(* IEC 61131-3 sources: volt/packages/volt-lsp-iec/test-corpus/pro2193/Device/Plc Logic/Application/09 Misc/Library Manager/CAA SegBufMan, 38 files *)

(* ---- ERROR.dut ---- *)
TYPE ERROR :
(
	NO_ERROR := 0,
	FIRST_ERROR := 6100,
	TIME_OUT,
	FIRST_MF,
	LAST_ERROR := 6199
);
END_TYPE

(* ---- RSHANDLING.gvl ---- *)
VAR_GLOBAL
	G_BUFFERCLASS : BufferClass;
	G_QUEUECLASS : QueueClass;
END_VAR

(* ---- VERSIONCONSTANTS.gvl ---- *)
VAR_GLOBAL
	GC_BYVERSION : BYTE := 1;
	GC_BYVERSION_1 : BYTE := 0;
END_VAR

(* ---- _BUFFERADDREF.pou ---- *)
FUNCTION _BUFFERADDREF : ERROR
VAR_INPUT
	HBUFFER : CAA.HANDLE;
END_VAR
END_FUNCTION

(* ---- _CHAINBUFFER.pou ---- *)
FUNCTION _CHAINBUFFER : CAA.HANDLE
VAR_INPUT
	HHEAD : CAA.HANDLE;
	HTAIL : CAA.HANDLE;
	PEERROR : POINTER TO ERROR;
END_VAR
END_FUNCTION

(* ---- _COPYBUFFERDATA.pou ---- *)
FUNCTION _COPYBUFFERDATA : ERROR
VAR_INPUT
	HBUFFER : CAA.HANDLE;
	SZOFFSET : CAA.SIZE;
	SZLENGTH : CAA.SIZE;
	PDATA : CAA.PVOID;
	SZSIZE : CAA.SIZE;
END_VAR
END_FUNCTION

(* ---- _CREATEBUFFER.pou ---- *)
FUNCTION _CREATEBUFFER : CAA.HANDLE
VAR_INPUT
	SZSIZE : CAA.SIZE;
	PDATA : CAA.PVOID;
	XPERMANENT : BOOL;
	PEERROR : POINTER TO ERROR;
END_VAR
END_FUNCTION

(* ---- _CREATEQUEUE.pou ---- *)
FUNCTION _CREATEQUEUE : CAA.HANDLE
VAR_INPUT
	PEERROR : POINTER TO ERROR;
END_VAR
END_FUNCTION

(* ---- _DELETEBUFFER.pou ---- *)
FUNCTION _DELETEBUFFER : ERROR
VAR_INPUT
	HBUFFER : CAA.HANDLE;
END_VAR
END_FUNCTION

(* ---- _DELETEQUEUE.pou ---- *)
FUNCTION _DELETEQUEUE : ERROR
VAR_INPUT
	HQUEUE : CAA.HANDLE;
END_VAR
END_FUNCTION

(* ---- _DEQUEUEBUFFER.pou ---- *)
FUNCTION _DEQUEUEBUFFER : CAA.HANDLE
VAR_INPUT
	HQUEUE : CAA.HANDLE;
	PEERROR : POINTER TO ERROR;
END_VAR
END_FUNCTION

(* ---- _ENQUEUEBUFFER.pou ---- *)
FUNCTION _ENQUEUEBUFFER : ERROR
VAR_INPUT
	HQUEUE : CAA.HANDLE;
	HBUFFER : CAA.HANDLE;
END_VAR
END_FUNCTION

(* ---- _GETBUFFERSIZE.pou ---- *)
FUNCTION _GETBUFFERSIZE : CAA.SIZE
VAR_INPUT
	HBUFFER : CAA.HANDLE;
	PEERROR : POINTER TO ERROR;
END_VAR
END_FUNCTION

(* ---- _GETQUEUELENGTH.pou ---- *)
FUNCTION _GETQUEUELENGTH : CAA.SIZE
VAR_INPUT
	HQUEUE : CAA.HANDLE;
	PEERROR : POINTER TO ERROR;
END_VAR
END_FUNCTION

(* ---- _GETSEGMENTDATAPOINTER.pou ---- *)
FUNCTION _GETSEGMENTDATAPOINTER : CAA.PVOID
VAR_INPUT
	HBUFFER : CAA.HANDLE;
	PSZSIZE : POINTER TO CAA.SIZE;
	PXPERMANENT : POINTER TO BOOL;
	PEERROR : POINTER TO ERROR;
END_VAR
END_FUNCTION

(* ---- _MOVETOBUFFEROFFSET.pou ---- *)
FUNCTION _MOVETOBUFFEROFFSET : ERROR
VAR_INPUT
	HBUFFER : CAA.HANDLE;
	SZOFFSET : CAA.SIZE;
END_VAR
END_FUNCTION

(* ---- _MOVETONEXTSEGMENT.pou ---- *)
FUNCTION _MOVETONEXTSEGMENT : ERROR
VAR_INPUT
	HBUFFER : CAA.HANDLE;
END_VAR
END_FUNCTION

(* ---- _SLICEBUFFER.pou ---- *)
FUNCTION _SLICEBUFFER : CAA.HANDLE
VAR_INPUT
	HBUFFER : CAA.HANDLE;
	SZOFFSET : CAA.SIZE;
	SZLENGTH : CAA.SIZE;
	PEERROR : POINTER TO ERROR;
END_VAR
END_FUNCTION

(* ---- CHAINBUFFER.pou ---- *)
FUNCTION CHAINBUFFER : CAA.HANDLE
VAR_INPUT
	HHEAD : CAA.HANDLE;
	HTAIL : CAA.HANDLE;
	PEERROR : POINTER TO ERROR;
END_VAR
END_FUNCTION

(* ---- COPYBUFFERDATA.pou ---- *)
FUNCTION COPYBUFFERDATA : ERROR
VAR_INPUT
	HBUFFER : CAA.HANDLE;
	SZOFFSET : CAA.SIZE;
	SZLENGTH : CAA.SIZE;
	PDATA : CAA.PVOID;
	SZSIZE : CAA.SIZE;
END_VAR
END_FUNCTION

(* ---- CREATEBUFFER.pou ---- *)
FUNCTION CREATEBUFFER : CAA.HANDLE
VAR_INPUT
	SZSIZE : CAA.SIZE;
	PDATA : CAA.PVOID;
	XPERMANENT : BOOL;
	PEERROR : POINTER TO ERROR;
END_VAR
END_FUNCTION

(* ---- CREATEQUEUE.pou ---- *)
FUNCTION CREATEQUEUE : CAA.HANDLE
VAR_INPUT
	PEERROR : POINTER TO ERROR;
END_VAR
END_FUNCTION

(* ---- DELETEBUFFER.pou ---- *)
FUNCTION DELETEBUFFER : ERROR
VAR_INPUT
	HBUFFER : CAA.HANDLE;
END_VAR
END_FUNCTION

(* ---- DELETEQUEUE.pou ---- *)
FUNCTION DELETEQUEUE : ERROR
VAR_INPUT
	HQUEUE : CAA.HANDLE;
END_VAR
END_FUNCTION

(* ---- DEQUEUEBUFFER.pou ---- *)
FUNCTION DEQUEUEBUFFER : CAA.HANDLE
VAR_INPUT
	HQUEUE : CAA.HANDLE;
	PEERROR : POINTER TO ERROR;
END_VAR
END_FUNCTION

(* ---- ENQUEUEBUFFER.pou ---- *)
FUNCTION ENQUEUEBUFFER : ERROR
VAR_INPUT
	HQUEUE : CAA.HANDLE;
	HBUFFER : CAA.HANDLE;
END_VAR
END_FUNCTION

(* ---- GETBUFFERSIZE.pou ---- *)
FUNCTION GETBUFFERSIZE : CAA.SIZE
VAR_INPUT
	HBUFFER : CAA.HANDLE;
	PEERROR : POINTER TO ERROR;
END_VAR
END_FUNCTION

(* ---- GETLIBVERSION.pou ---- *)
FUNCTION GETLIBVERSION : VERSION
END_FUNCTION

(* ---- GETLIBVERSIONNUMBER.pou ---- *)
FUNCTION GETLIBVERSIONNUMBER : DWORD
END_FUNCTION

(* ---- GETQUEUELENGTH.pou ---- *)
FUNCTION GETQUEUELENGTH : CAA.SIZE
VAR_INPUT
	HQUEUE : CAA.HANDLE;
	PEERROR : POINTER TO ERROR;
END_VAR
END_FUNCTION

(* ---- GETSEGMENTDATAPOINTER.pou ---- *)
FUNCTION GETSEGMENTDATAPOINTER : CAA.PVOID
VAR_INPUT
	HBUFFER : CAA.HANDLE;
	PSZSIZE : POINTER TO CAA.SIZE;
	PXPERMANENT : POINTER TO BOOL;
	PEERROR : POINTER TO ERROR;
END_VAR
END_FUNCTION

(* ---- GETSUPPLIERVERSION.pou ---- *)
FUNCTION GETSUPPLIERVERSION : WORD
VAR_INPUT
	XDUMMY : BOOL;
END_VAR
END_FUNCTION

(* ---- ISLIBRELEASED.pou ---- *)
FUNCTION ISLIBRELEASED : BOOL
END_FUNCTION

(* ---- MOVETOBUFFEROFFSET.pou ---- *)
FUNCTION MOVETOBUFFEROFFSET : ERROR
VAR_INPUT
	HBUFFER : CAA.HANDLE;
	SZOFFSET : CAA.SIZE;
END_VAR
END_FUNCTION

(* ---- MOVETONEXTSEGMENT.pou ---- *)
FUNCTION MOVETONEXTSEGMENT : ERROR
VAR_INPUT
	HBUFFER : CAA.HANDLE;
END_VAR
END_FUNCTION

(* ---- SLICEBUFFER.pou ---- *)
FUNCTION SLICEBUFFER : CAA.HANDLE
VAR_INPUT
	HBUFFER : CAA.HANDLE;
	SZOFFSET : CAA.SIZE;
	SZLENGTH : CAA.SIZE;
	PEERROR : POINTER TO ERROR;
END_VAR
END_FUNCTION

(* ---- BUFFERCLASS.pou ---- *)
FUNCTION_BLOCK BUFFERCLASS EXTENDS RSMClass
END_FUNCTION_BLOCK

METHOD CLOSE : RSM.ERROR
VAR_INPUT
	HHANDLE : CAA.HANDLE;
END_VAR
END_METHOD

(* ---- QUEUECLASS.pou ---- *)
FUNCTION_BLOCK QUEUECLASS EXTENDS RSMClass
END_FUNCTION_BLOCK

METHOD CLOSE : RSM.ERROR
VAR_INPUT
	HHANDLE : CAA.HANDLE;
END_VAR
END_METHOD
